(* IEC 61131-3 sources: traffic-lights/PLC_TrafficLights/Class/Varan_Base (part 2) *)

  ud_timeout := ud_ResponseTimeMax + ud_bytes * VM_TIMEOUT_ONE_BYTE + VM_RETRY_TIMEOUT_STD_OFFSET;

END_FUNCTION // Varan_Base::GetRetryTimeout
//=================================================================================================
//---------------------- Additional functions------------------------------------------------------
//=================================================================================================

//[#ENGLISH]
//=================================================================================================
//Function to Start time measurement
//=================================================================================================
#pragma warning(disable:74)
#pragma warning(disable:73)
FUNCTION Varan_Base::StartTimeMeasurement
  VAR_INPUT
    usMode (EAX) 	: DINT;
  END_VAR
#ifdef VM_CLASS_TIME_MEASUREMENT
  VAR
    tmpTime : ^t_TimeMeasurementVaran;
  END_VAR

  case usMode of

    //-----------------------------------------------------------

    VARANTIME_RT:
      tmpTime := #s_TimeRt;

    //-----------------------------------------------------------

    VARANTIME_RTPOSTSCAN:
      tmpTime := #s_TimeRtPostScan;

    //-----------------------------------------------------------

    VARANTIME_CY:
      tmpTime := #s_TimeCy;

    //-----------------------------------------------------------

  end_case;

  if ( tmpTime^.us_Activate ) then
    tmpTime^.ud_Timemark := VaranIn.GetNsTime();
  end_if;

#endif

END_FUNCTION // Varan_Base::StartTimeMeasurement
//[#ENGLISH]
//=================================================================================================
//Function to Stop time measurement
//=================================================================================================
FUNCTION Varan_Base::StopTimeMeasurement
  VAR_INPUT
    usMode (EAX) 	: DINT;
  END_VAR
#ifdef VM_CLASS_TIME_MEASUREMENT
  VAR
    tmpTime : ^t_TimeMeasurementVaran;
  END_VAR

  case usMode of

    //-----------------------------------------------------------

    VARANTIME_RT:
      tmpTime := #s_TimeRt;

    //-----------------------------------------------------------

    VARANTIME_RTPOSTSCAN:
      tmpTime := #s_TimeRtPostScan;

    //-----------------------------------------------------------

    VARANTIME_CY:
      tmpTime := #s_TimeCy;

    //-----------------------------------------------------------

  end_case;

  if ( tmpTime^.us_Activate ) then

    //get actual time
    tmpTime^.ud_ActualTime := VaranIn.GetNsTime() - tmpTime^.ud_Timemark;

    //look for maximum time
    if ( tmpTime^.ud_ActualTime > tmpTime^.ud_MaximalTime ) then
      tmpTime^.ud_MaximalTime := tmpTime^.ud_ActualTime;
    end_if;

    //look for minimum time
    if ( tmpTime^.ud_ActualTime < tmpTime^.ud_MinimalTime ) then
      tmpTime^.ud_MinimalTime := tmpTime^.ud_ActualTime;
    end_if;

    //look for average time (100000 cycles)
    if ( tmpTime^.ud_AverageCounter = 100000 ) then

      tmpTime^.ud_AverageTime 	:= tmpTime^.ud_AverageSum / tmpTime^.ud_AverageCounter;
      tmpTime^.ud_AverageSum 	:= 0;
      tmpTime^.ud_AverageCounter := 0;

    else
      tmpTime^.ud_AverageSum += ( tmpTime^.ud_ActualTime / 100 );
      tmpTime^.ud_AverageCounter += 1;
    end_if;
  end_if;

#endif

END_FUNCTION // Varan_Base::StopTimeMeasurement
#pragma warning(default:74)
#pragma warning(default:73)

//[#ENGLISH]
//=================================================================================================
//Function to set state of class
//=================================================================================================
//[>sd_error]type of error
FUNCTION VIRTUAL GLOBAL Varan_Base::SetState
  VAR_INPUT
    sd_error		: t_e_VaranErrors;
  END_VAR

  //only set error if class is ok
  if ( State = _ClassOk ) then

    State := sd_error;

  else
    //only eeprom error can be cleared
    if ( State = _EEPromError & sd_error = _ClassOk ) then
      State := sd_error;
    end_if;
  end_if;

END_FUNCTION //VIRTUAL GLOBAL Varan_Base::SetState
//[#ENGLISH]
//=================================================================================================
//Function to disable device
//=================================================================================================
//[<sd_retval]0=ok, -17=Port no link, -30=client disabled, -31=client cant enable, -100 function not available with this os version, other return code of os
FUNCTION VIRTUAL GLOBAL Varan_Base::DisableDevice
  VAR_OUTPUT
    sd_retval	: DINT;
  END_VAR
  VAR
    nodeProperty    : LSL_PROPERTY_VALUE_PAIR;
  END_VAR

  //look if funtion is available with this os version
  if ( _RTOSVersion >= VM_DISABLE_DEVICE_AVAILABLE ) then

    if b_PayloadSupport then
      nodeProperty.udPropertyId    := ND_PROP_CONNECTION_STATE;
      nodeProperty.udPropertyValue := CN_STATE_DISCONNECTED;
      sd_retval := MULTI_VARAN_iSetNodeProperties(  hNodeHandle           := ud_HandleModule
                                                  , udPropertyCount       := 1
                                                  , psPropertyValuePairs  := #nodeProperty);
    else
      //disable device
      sd_retval := VARAN_iSetNodeEnableStatus	( uiManager		:= ud_VaranManagerNr
                          , pucNode		:= p_VaranPosition
                          , uiNodeStatus	:= 0
                          );
    end_if;

    // if there was an error at disabling it was not caused by a disabled previous module
    if	( sd_retval <> VARANMANAGER_OK ) &
        ( sd_retval <> VARANMANAGER_CLIENT_DISABLED ) &
        ( sd_retval <> VARANMANAGER_ADMIN_DOL_EXECUTION_ERROR	) &	//because if device before is disabled, DA can't work
        ( VaranIn.IsDeviceDisabled() = FALSE ) then

      State := _DisableError;

      //Set VaranMaster off
      VaranIn.SetManagerOff( e_error := State );
    end_if;

    //port is disabled
    b_DisableDevice := FALSE;
    ud_DisableTime := ops.tAbsolute;
  else
    b_DisableDevice := FALSE;
    sd_retval := -100;
  end_if;

  // Force end of Cylic Post Init
  if bPostInitNeeded then
    CheckCyclicPostInitFinished(TRUE);
  end_if;

END_FUNCTION // Varan_Base::DisableDevice
//[#ENGLISH]
//=================================================================================================
//Function to enable device
//=================================================================================================
//[<sd_retval]0=ok, 1=device must disabled for more then 200ms, 2=-100 function not available with this os version, -17=Port no link, -30=client disabled, -31=client cant enable, other return code of os
FUNCTION VIRTUAL GLOBAL Varan_Base::EnableDevice
  VAR_OUTPUT
    sd_retval	: DINT;
  END_VAR
  VAR
    nodeProperty    : LSL_PROPERTY_VALUE_PAIR;
  END_VAR

  //look if funtion is available with this os
  if ( _RTOSVersion >= VM_DISABLE_DEVICE_AVAILABLE ) then

    //look if watchdog time is gone
    if ( ( ops.tAbsolute - ud_DisableTime ) < 200ms ) then
      sd_retval := 1;
      return;
    end_if;

    if b_PayloadSupport then
      nodeProperty.udPropertyId    := ND_PROP_CONNECTION_STATE;
      nodeProperty.udPropertyValue := CN_STATE_CONNECTED;
      sd_retval := MULTI_VARAN_iSetNodeProperties(  hNodeHandle           := ud_HandleModule
                                                  , udPropertyCount       := 1
                                                  , psPropertyValuePairs  := #nodeProperty);
    else
      //enable device
      sd_retval := VARAN_iSetNodeEnableStatus	( uiManager		:= ud_VaranManagerNr
                          , pucNode		:= p_VaranPosition
                          , uiNodeStatus	:= 1
                          );
    end_if;

    //look for an error
    if ( sd_retval <> VARANMANAGER_OK ) then
      State := _EnableError;
    end_if;
  else
    sd_retval := 2;
  end_if;

END_FUNCTION // Varan_Base::EnableDevice
//[#ENGLISH]
//=================================================================================================
//Function to set all Data Objects off
//=================================================================================================
FUNCTION VIRTUAL GLOBAL Varan_Base::SetDOsOff

  //in base class we have no DO's

END_FUNCTION // Varan_Base::SetDOsOff
//[#ENGLISH]
//=================================================================================================
//Function to look if class is disabled
//=================================================================================================
//[<b_disabled]TRUE -> Device is disabled
FUNCTION VIRTUAL GLOBAL Varan_Base::IsDeviceDisabled
  VAR_OUTPUT
    b_disabled		: BOOL;
  END_VAR

  if 	( State = _NoHardware
    | State = _HardwareNotRequiredIRQ
    )
  then
    b_disabled := TRUE;
  else
    //look class above
    b_disabled := VaranIn.IsDeviceDisabled();
  end_if;

END_FUNCTION //VIRTUAL GLOBAL Varan_Base::IsDeviceDisabled
//[#ENGLISH]
//=================================================================================================
//Function to set multiple memory read/write options
//=================================================================================================
//[>us_filter]filter of multicast write
//[>us_sequence]sequence number of device
//[<sd_retval]error code
FUNCTION VIRTUAL GLOBAL Varan_Base::SetMultipleSettings
  VAR_INPUT
    us_filter		: USINT;
    us_sequence		: usint;
  END_VAR
  VAR_OUTPUT
    sd_retval		: DINT;
  END_VAR
  VAR
    a_data			: ARRAY[0..10] OF USINT;
  END_VAR

  //look if class is ok
  if ( State = _ClassOk ) then

    us_MulticastFilter 		:= us_filter;
    us_MultipleSequence		:= us_sequence;

    //set data for direct access
    a_data[ 0 ] := us_MulticastFilter;
    a_data[ 3 ] := us_sequence;
    a_data[ 10 ] := 16#6;					//to trigger watchdog only with watchdog command and multiple read/write command

    // Payload Support
    if b_PayloadSupport then
      //write data with direct access
      sd_retval := MULTI_VARAN_iExecuteDirectAccess(  hNodeHandle := ud_HandleModule
                                                    , udCommand   := VARAN_CMD_CONTROL_WRITE
                                                    , udOffset    := VARAN_MULTIPLE_OFFSET
                                                    , udLength    := sizeof(a_data)
                                                    , pusData     := ( #a_data )$^USINT
                                                    , pudErrorInfo:= NIL);
    else
      //write data with direct access
      sd_retval := VARAN_iWriteControlDA	( uiManager		  := ud_VaranManagerNr
                                          , uiAddress		  := DeviceAddress + VARAN_MULTIPLE_OFFSET
                                          , uiLen			    := sizeof(a_data)
                                          , uiRetryTimeout:= GetRetryTimeout( ud_bytes := sizeof(a_data) )
                                          , pvData		    := ( #a_data )$^UDINT
                                          , puiError		  := NIL
                                          );
    end_if;

    //look if an error occurs
    if ( sd_retval <> VARANMANAGER_OK ) then
      State := _MultipleError;
      return;
    end_if;
  end_if;

END_FUNCTION //VIRTUAL GLOBAL Varan_Base::SetMultipleSettings
//[#ENGLISH]
//=================================================================================================
//Function must be overwrite
//=================================================================================================
//[>p_handle]pointer to data object header
//[>p_data_read]pointer to read data
//[>p_data_write]pointer to data write
//[<sd_retval]error code
#pragma warning(disable: 73)
FUNCTION VIRTUAL GLOBAL Varan_Base::SetMultipleDataPointers
  VAR_INPUT
    p_handle		: ^LSL_VARANFRAME;
    p_data_read		: ^UDINT;
    p_data_write	: ^UDINT;
    DOIndex         : UDINT;
  END_VAR
  VAR_OUTPUT
    sd_retval		: DINT;
  END_VAR

  sd_retval := -1;

END_FUNCTION //VIRTUAL GLOBAL Varan_Base::SetMultipleDataPointers
#pragma warning(default: 73)
//[#ENGLISH]
//=================================================================================================
//Function to get pointer to calib data
//=================================================================================================
//[>p_offset]pointer to variable to write offset
//[<sd_retval]errorcode of os
FUNCTION  Varan_Base::GetCalibDataPointer
  VAR_INPUT
    p_offset	: ^UDINT;
  END_VAR
  VAR_OUTPUT
    sd_retval	: DINT;
  END_VAR
  VAR
    a_data			: ARRAY[0..31] OF UDINT;
    i				: UDINT;
  END_VAR

  //read SPI data
  sd_retval := VaranIn.ReadSPIData( p_us_position_info	:= p_VaranPosition
                  , ud_offset				:= 0
                  , ud_length				:= 128 or VM_SPI_IDENT_LIST
                  , p_data				:= ( #a_data )$^USINT
                  );

  //look for an error
  if ( sd_retval <> VARANMANAGER_OK ) then
    State := _SPIError;
    return;
  end_if;

  //look for right Identifier
  if ( a_data[ 0 ] <> 16#12345678 ) then
    State := _SPIError;
    return;
  end_if;

  //look for valid length	(we only read 128 Byte at the moment [16Byte are header])
  if( a_data[ 3 ] > (128 - 16 ) ) then
    State := _SPIError;
    return;
  end_if;

  //search for calib data
  for i := 0 to a_data[ 3 ] / sizeof( UDINT ) do

    //look for calib id in 3rd byte
    if ( ( a_data[ i + 4 ] and 16#FF00_0000 ) = VM_SPI_CALIB_ID ) then
      p_offset^ := a_data[ i + 4 ] and 16#00FF_FFFF;
      return;
    end_if;
  end_for;

  //if no entry is found
  State := _NoCalibDataFound;
  sd_retval := -100;

END_FUNCTION // Varan_Base::GetCalibDataPointer
//[#ENGLISH]
//=================================================================================================
//Function to get pointer to calib data
//=================================================================================================
//[>ud_offset]offset in SPI - Flash
//[>ud_length]length of data
//[>p_data]pointer to allocated data space
//[<sd_retval]return value of OS
FUNCTION  Varan_Base::ReadSPIData
  VAR_INPUT
    ud_offset	: UDINT;
    ud_length	: UDINT;
    p_data		: ^USINT;
  END_VAR
  VAR_OUTPUT
    sd_retval	: DINT;
  END_VAR
  VAR
    ud_read_length	: UDINT;
  END_VAR

  //look if we have a length
  if ( ud_length = 0 ) then
    sd_retval := -100;
    return;
  end_if;

  //look if data is in one page
  while ( ud_length <> 0 ) do

    //if length is above page size
    if ( ( ud_offset and 16#FF ) + ud_length > 16#FF ) then
      //how many bytes are in this page available
      ud_read_length := 16#100 - ( ud_offset and 16#FF );
      //not more than 128 Bytes
      if ( ud_read_length > 128 ) then
        ud_read_length := 128;
      end_if;
    else
      //not more than 128 Bytes
      if ( ud_length > 128 ) then
        ud_read_length := 128;
      else
        ud_read_length := ud_length;
      end_if;
    end_if;

    //read data
    sd_retval := VaranIn.ReadSPIData( p_us_position_info	:= p_VaranPosition
                    , ud_offset				:= ud_offset
                    , ud_length				:= ud_read_length
                    , p_data				:= p_data
                    );
    //look for an error
    if ( sd_retval <> VARANMANAGER_OK ) then
      State := _SPIError;
      return;
    end_if;

    //correct length
    ud_length -= ud_read_length;
    ud_offset += ud_read_length;
    p_data += ud_read_length;
  end_while;

END_FUNCTION // Varan_Base::ReadSPIData

//[#ENGLISH]
//=================================================================================================
//Function to update module retry counter
//=================================================================================================
FUNCTION VIRTUAL GLOBAL Varan_Base::UpdateRetryCounter
  //function must be override
END_FUNCTION //VIRTUAL GLOBAL Varan_Base::UpdateRetryCounter
//[#ENGLISH]
//=================================================================================================
//Function to get varan time
//=================================================================================================
//[<ud_varan_time]varan time
FUNCTION VIRTUAL GLOBAL Varan_Base::GetVaranTime
  VAR_INPUT
    p_ud_IsoStartPoint	: ^UDINT;
  END_VAR
  VAR_OUTPUT
    ud_varan_time		: UDINT;
  END_VAR

  ud_varan_time := VaranIn.GetVaranTime( p_ud_IsoStartPoint );

END_FUNCTION //VIRTUAL GLOBAL Varan_Base::GetVaranTime
//[#ENGLISH]
//=================================================================================================
//Function to disable Device in Rt (because VARAN_iSetNodeEnableStatus must not called in Realtime)
//=================================================================================================
FUNCTION  Varan_Base::DisableDeviceRt
  VAR_OUTPUT
    sd_retval		: DINT;
  END_VAR

  //look if funtion is available with this os version
  if ( _RTOSVersion >= VM_DISABLE_DEVICE_AVAILABLE ) then

      //disable device
    sd_retval := VaranIn.SetDisableDevice( p_us_position_info := p_VaranPosition );

    //check error
      if ( sd_retval = 0 ) then

        //port is disabled
        b_DisableDevice := FALSE;
        ud_DisableTime := ops.tAbsolute;
      end_if;
  else
    b_DisableDevice := FALSE;
    sd_retval := -100;
  end_if;

  // Force end of Cylic Post Init
  if bPostInitNeeded then
    CheckCyclicPostInitFinished(TRUE);
  end_if;

END_FUNCTION // Varan_Base::DisableDeviceRt

FUNCTION Varan_Base::SetNewPllData
  VAR_INPUT
    ud_delay_time 	: UDINT;
    us_divider 	    : USINT;
  END_VAR
  VAR_OUTPUT
    sd_retval 	    : DINT;
  END_VAR
  VAR
    ud_data			    : UDINT;
  END_VAR

  //calculate right register value (Response Time (in 10ns steps) / 2 - constant FPGA delay time
  ud_DeviceDelayTime := ( p_NodeInfo^.uiResponseTime ) / 20 + VM_CONST_FPGA_DELAY + ud_delay_time;

  // Payload support
  if b_PayloadSupport then
    //write Pll time with direct access
    sd_retval := MULTI_VARAN_iExecuteDirectAccess(  hNodeHandle := ud_HandleModule
                                                  , udCommand   := VARAN_CMD_CONTROL_WRITE
                                                  , udOffset    := VARAN_PLL_OFFSET + 16#C
                                                  , udLength    := 3
                                                  , pusData     := ( #ud_DeviceDelayTime )$^USINT
                                                  , pudErrorInfo:= NIL);
  else
    //write Pll time with direct access
    sd_retval := VARAN_iWriteControlDA( uiManager		  := ud_VaranManagerNr
                                      , uiAddress		  := DeviceAddress + VARAN_PLL_OFFSET + 16#C
                                      , uiLen			    := 3
                                      , uiRetryTimeout:= GetRetryTimeout( ud_bytes := 3 )
                                      , pvData		    := ( #ud_DeviceDelayTime )$^UDINT
                                      , puiError		  := NIL
                                      );
  end_if;

  //look if an error occurs
  if ( sd_retval <> VARANMANAGER_OK ) then
    State := _PllError;
    return;
  end_if;

  //set divider (only for new pll if function is available)
  if ( us_divider <> 0 ) then

    if b_PayloadSupport then  //  -------------------------------------------------------------------------
      // disable divider
      ud_data := 0;

      sd_retval := MULTI_VARAN_iExecuteDirectAccess(  hNodeHandle := ud_HandleModule
                                                    , udCommand   := VARAN_CMD_CONTROL_WRITE
                                                    , udOffset    := VARAN_PLL_OFFSET + 16#A
                                                    , udLength    := 1
                                                    , pusData     := ( #ud_data )$^USINT
                                                    , pudErrorInfo:= NIL);

      //look if an error occurs
      if ( sd_retval <> VARANMANAGER_OK ) then
        State := _PllError;
        return;
      end_if;

      // set divider value
      ud_data := us_divider;

      sd_retval := MULTI_VARAN_iExecuteDirectAccess(  hNodeHandle := ud_HandleModule
                                                    , udCommand   := VARAN_CMD_CONTROL_WRITE
                                                    , udOffset    := VARAN_PLL_OFFSET + 16#B
                                                    , udLength    := 1
                                                    , pusData     := ( #ud_data )$^USINT
                                                    , pudErrorInfo:= NIL);

      //look if an error occurs
      if ( sd_retval <> VARANMANAGER_OK ) then
        State := _PllError;
        return;
      end_if;

      // enable divider
      ud_data := 2#10010000;    //Defaultvalue = 0x80 + SyncDivider Eanble Bit (Bit4)

      sd_retval := MULTI_VARAN_iExecuteDirectAccess(  hNodeHandle := ud_HandleModule
                                                    , udCommand   := VARAN_CMD_CONTROL_WRITE
                                                    , udOffset    := VARAN_PLL_OFFSET + 16#A
                                                    , udLength    := 1
                                                    , pusData     := ( #ud_data )$^USINT
                                                    , pudErrorInfo:= NIL);

      //look if an error occurs
      if ( sd_retval <> VARANMANAGER_OK ) then
        State := _PllError;
        return;
      end_if;

    else  // if b_PayloadSupport -------------------------------------------------------------------------

      // disable divider
      ud_data := 0;

      // write control register
      sd_retval := VARAN_iWriteControlDA( uiManager		  := ud_VaranManagerNr
                                        , uiAddress		  := DeviceAddress + VARAN_PLL_OFFSET + 16#A
                                        , uiLen			    := 1
                                        , uiRetryTimeout:= GetRetryTimeout( ud_bytes := 1 )
                                        , pvData		    := ( #ud_data )$^UDINT
                                        , puiError		  := NIL
                                        );

      //look if an error occurs
      if ( sd_retval <> VARANMANAGER_OK ) then
        State := _PllError;
        return;
      end_if;

      // set divider value
      ud_data := us_divider;

      //write Divider with direct access
      sd_retval := VARAN_iWriteControlDA( uiManager		  := ud_VaranManagerNr
                                        , uiAddress		  := DeviceAddress + VARAN_PLL_OFFSET + 16#B
                                        , uiLen			    := 1
                                        , uiRetryTimeout:= GetRetryTimeout( ud_bytes := 1 )
                                        , pvData		    := ( #ud_data )$^UDINT
                                        , puiError		  := NIL
                                        );

      //look if an error occurs
      if ( sd_retval <> VARANMANAGER_OK ) then
        State := _PllError;
        return;
      end_if;

      // enable divider
      ud_data := 2#10010000;    //Defaultvalue = 0x80 + SyncDivider Eanble Bit (Bit4)

      //write Divider with direct access
      sd_retval := VARAN_iWriteControlDA( uiManager		  := ud_VaranManagerNr
                                        , uiAddress		  := DeviceAddress + VARAN_PLL_OFFSET + 16#A
                                        , uiLen			    := 1
                                        , uiRetryTimeout:= GetRetryTimeout( ud_bytes := 1 )
                                        , pvData		    := ( #ud_data )$^UDINT
                                        , puiError		  := NIL
                                        );

      //look if an error occurs
      if ( sd_retval <> VARANMANAGER_OK ) then
        State := _PllError;
        return;
      end_if;

    end_if; // if b_PayloadSupport -------------------------------------------------------------------------

  end_if; // us_divider <> 0

END_FUNCTION

FUNCTION VIRTUAL GLOBAL Varan_Base::GetDocumentation
  VAR_INPUT
    p_dpne 	: ^CHAR;
  END_VAR
  VAR_OUTPUT
    sd_retval 	: DINT;
  END_VAR

  sd_retval := VaranIn.GetDocumentation(p_us_position_info:=p_VaranPosition, p_dpne:=p_dpne);

END_FUNCTION

FUNCTION VIRTUAL GLOBAL Varan_Base::UpdateRtPostScan

END_FUNCTION

FUNCTION GLOBAL Varan_Base::SetRunStatus
  VAR_INPUT
    state 	: USINT;
  END_VAR
  VAR_OUTPUT
    us_retval 	: USINT;
  END_VAR

  if Required then
    us_retval := state or VARAN_DO_REQUIRED;
  else
    us_retval := state;
  end_if;

END_FUNCTION

FUNCTION VIRTUAL GLOBAL Varan_Base::GetPointer2ObjectPath
  VAR_OUTPUT
    p_us_ObjectPath 	: ^USINT;
  END_VAR
  VAR
    i                       : USINT;
    udSystemVaranManagerCnt : UDINT;
    _Para 	                : CmdStruct;
    _Result 	              : Results;
  END_VAR

  if ( p_ObjectPath = NIL ) then

    if ( p_VaranPosition = NIL ) then

      Varan_Base::Init();

      if ( p_VaranPosition = NIL ) then

        p_us_ObjectPath := NIL;
        return;

      end_if;
    end_if;

    if ( p_VaranPosition^ >= VARAN_MAX_DEPTH ) then
      p_us_ObjectPath := NIL;
      return;
    end_if;

    //alloc memory
    p_ObjectPath := ( To_StdLib.Malloc( size := p_VaranPosition^ + 5 ) )$^USINT;

    To_StdLib.MemCpy( dest 		:= p_ObjectPath
                    , source	:= p_VaranPosition
                    , size		:= p_VaranPosition^ + 1
                    );

    _Para.uiCmd := VM_CMD_GET_SYSTEM_MANAGER_CNT;
    _Result.aData[0]$UDINT  := 1;   // Set to 1 in case the NewInst Method is not Implemented
    udSystemVaranManagerCnt := 1;

    if VaranIn.NewInst(#_Para, #_Result) = READY then
      udSystemVaranManagerCnt := _Result.aData[0]$UDINT;
    end_if;

    //Check if we have to build the "new" hardware tree with the new escape sequence
    if udSystemVaranManagerCnt > 1 then

      //More than one manager --> new HW-Tree with new esacpe sequence

      //insert one byte after length
      for i := p_ObjectPath^ to 1 by -1 do
        ( p_ObjectPath + i + 4 )^ := ( p_ObjectPath + i )^;
      end_for;

      // domain info byte
      ( p_ObjectPath + 1 )^ := 0;

      //insert escape sequence for varan
      ( p_ObjectPath + 2 )^ := HWT_ESCAPE_MULTIVARAN;

      //insert escape sequence for varan
      ( p_ObjectPath + 3 )^ := ud_VaranManagerNr$USINT;

      //insert escape sequence for varan
      ( p_ObjectPath + 4 )^ := HWT_ESCAPE_VARAN;

      //increase length
      p_ObjectPath^ += 4;

    else

      //Old HW-Tree (without Multivaran Escape sequence)

      //insert one byte after length
      for i := p_ObjectPath^ to 1 by -1 do
        ( p_ObjectPath + i + 2 )^ := ( p_ObjectPath + i )^;
      end_for;

      // domain info byte
      ( p_ObjectPath + 1 )^ := 0;

      //insert escape sequence for varan
      ( p_ObjectPath + 2 )^ := HWT_ESCAPE_VARAN;

      //increase length
      p_ObjectPath^ += 2;

    end_if;

    //register object path in OS
    SetObjectThisp(p_us_ObjectPath:=p_ObjectPath, ud_thisp:=this$UDINT);

  end_if;

  p_us_ObjectPath := p_ObjectPath;

END_FUNCTION

FUNCTION VIRTUAL GLOBAL Varan_Base::SetObjectThisp
  VAR_INPUT
    p_us_ObjectPath 	: ^USINT;
    ud_thisp 	: UDINT;
  END_VAR
  VAR_OUTPUT
    sd_retval 	: DINT;
  END_VAR

  sd_retval := VaranIn.SetObjectThisp(p_us_ObjectPath,ud_thisp);

END_FUNCTION

FUNCTION VIRTUAL GLOBAL Varan_Base::GetObjectThisp
  VAR_INPUT
    p_us_ObjectPath : ^USINT;
  END_VAR
  VAR_OUTPUT
    ud_Thisp 	      : UDINT;
  END_VAR

  ud_thisp := VaranIn.GetObjectThisp(p_us_ObjectPath:=p_us_ObjectPath);

END_FUNCTION

FUNCTION Varan_Base::Diagnose
#ifdef VARAN_DIAGNOSE
  VAR
    os_retcode : DINT;
  END_VAR

  if State = _ClassOk then
    os_retcode := VARAN_IGETVARANDIAGNOSTICS(8, #s_Diagnose.cmd_Input, s_Diagnose.InputSize, #s_Diagnose.cmd_Output, #s_Diagnose.OutputSize);

    //reset counter
    if s_Diagnose.Command = Reset then
      ConnectCounter      := 0;
      FaultCounter        := 0;
      RXLost              := 0;
      TXLost              := 0;
      s_Diagnose.Command  := Activate;
    end_if;

    //OS doesn't support Diagnose
    if os_retcode <> 0 then
      DiagControl := -1;
      return;
    end_if;

    //FPGA doesn't support Diagnose
    if s_Diagnose.cmd_Output.Flags.1 = 0 then
      DiagControl := -2;
      return;
    end_if;

    DiagControl     := 1;
    ConnectCounter  += s_Diagnose.cmd_Output.Counter1 - s_Diagnose.OldCounter.Counter1;
    FaultCounter    += s_Diagnose.cmd_Output.Counter2 - s_Diagnose.OldCounter.Counter2;
    RXLost          += s_Diagnose.cmd_Output.Counter3 - s_Diagnose.OldCounter.Counter3;
    TXLost          += s_Diagnose.cmd_Output.Counter4 - s_Diagnose.OldCounter.Counter4;

    s_Diagnose.OldCounter.Counter1 := s_Diagnose.cmd_Output.Counter1;
    s_Diagnose.OldCounter.Counter2 := s_Diagnose.cmd_Output.Counter2;
    s_Diagnose.OldCounter.Counter3 := s_Diagnose.cmd_Output.Counter3;
    s_Diagnose.OldCounter.Counter4 := s_Diagnose.cmd_Output.Counter4;
  end_if;
#endif
END_FUNCTION

#pragma warning(disable:73)
#pragma warning(disable:74)
#pragma warning(disable:76)
FUNCTION VIRTUAL GLOBAL Varan_Base::DiagControl::Write
  VAR_INPUT
    input (EAX) 	: DINT;
  END_VAR
  VAR_OUTPUT
    result (EAX) 	: DINT;
  END_VAR

#ifdef VARAN_DIAGNOSE

  if input >= 0 & input <= 2 then
    s_Diagnose.Command$DINT := input;
  end_if;

#endif

END_FUNCTION
#pragma warning(default:73)
#pragma warning(default:74)
#pragma warning(default:76)

FUNCTION VIRTUAL GLOBAL Varan_Base::ValidateSerNo::Write
  VAR_INPUT
    input (EAX) 	: DINT;
  END_VAR
  VAR_OUTPUT
    result (EAX) 	: DINT;
  END_VAR

  result := input;

  if (b_ValidationInProgress = FALSE) & SerNoValidation then

    To_MultiTask.CREATETHREAD(taskfunction0:=#SerNoValidationTask(),
                              priority0:=14,
                              stackSize0:=16#4000,
                              flags0:=MT_TASK_SAVETHIS,
                              parameter0:=this,
                              name0:=#szSerNoStr[0]);

    b_ValidationInProgress := TRUE;
  end_if;

END_FUNCTION

FUNCTION Varan_Base::SerNoValidationTask

  // get length of string
  SerNoHeader.StringLength := _strlen(#szSerNoStr[0]);

  // reserve enough space in ramfile
  if SerNoBackup.SetSize(sizeof(SerNoHeader) + SerNoHeader.StringLength) <> C_OK then
      b_ValidationInProgress := FALSE;
      return;
    end_if;

  // initialize the rest of the header
  SerNoHeader.Version := SERNO_VALIDATION_VERSION;
  SerNoHeader.ZeroByte := 0;

  // write to ramfile
  if (SerNoBackup.SetDataAt((#SerNoHeader)$^USINT, sizeof(SerNoHeader), 0) = C_OK) &
     (SerNoBackup.SetDataAt((#szSerNoStr[0])$^USINT, _strlen(#szSerNoStr[0]), sizeof(SerNoHeader)) = C_OK) then
    // if we had a problem with serial number before
    if State = _InvalidSerialNo then
      // try to reconnect
      Varan_HwConnect(0);
    end_if;

    ValidateSerNo := 1;
  else
    ValidateSerNo := 0;
  end_if;

  b_ValidationInProgress := FALSE;

END_FUNCTION

#pragma warning(disable:73)
FUNCTION VIRTUAL GLOBAL Varan_Base::CheckDeviceID
  VAR_INPUT
    ID2Check 	: UDINT;
  END_VAR
  VAR_OUTPUT
    IsOK 	: BOOL;
  END_VAR
#pragma warning(default:73)

  IsOK := TRUE;

END_FUNCTION

FUNCTION GLOBAL Varan_Base::FlexInit
  VAR
    sd_retval	: DINT;
  END_VAR

  //look for an error
  if ( pVaran = NIL ) then
    State := _NoVaranInterface;
    if Required then
      VaranIn.AllowRequiredError();
    end_if;
    return;
  end_if;

  //-----------------------------------------------------------------------------------------------
  //get Varan position if we have no position yet
  if ( p_VaranPosition = NIL ) then

    //alloc memory to get position
    p_VaranPosition := ( To_StdLib.Malloc( size := VARAN_MAX_DEPTH + 1 ) )$^USINT;
    //look if an error occurs
    if ( p_VaranPosition = NIL ) then
      State := _RootError;
      return;
    end_if;

  else

    //alloc memory for position pointer
    p_VaranPosition := 	( To_StdLib.ReAlloc	( mptr := p_VaranPosition , newsize	:= VARAN_MAX_DEPTH + 1))$^USINT;
    //look if an error occurs
    if ( p_VaranPosition = NIL ) then
      State := _RootError;
      return;
    end_if;

  end_if;

  //set length to 0
  p_VaranPosition^ := 0;

  //get position
  sd_retval := VaranIn.GetVaranPosition( p_us_info := p_VaranPosition );

  //look if an error occurs
  if ( sd_retval <> VARANMANAGER_OK ) then
    State := _RootError;
    return;
  end_if;

  //alloc memory for position pointer
  p_VaranPosition := 	( To_StdLib.ReAlloc	( mptr		:= p_VaranPosition
                      , newsize	:= p_VaranPosition^ + 1
                      )
            )$^USINT;

  //look if an error occurs
  if ( p_VaranPosition = NIL ) then
    State := _RootError;
    return;
  end_if;

  //-----------------------------------------------------------------------------------------------
  //install callback function
  sd_retval := InstallCallbackObject();

  //look if an error occurs
  if ( sd_retval <> VARANMANAGER_OK ) then
    State := _CallBackError;
    return;
  end_if;

END_FUNCTION

FUNCTION GLOBAL Varan_Base::AllowRequiredError

  VaranIn.AllowRequiredError();

END_FUNCTION

FUNCTION GLOBAL Varan_Base::IsTransparent
  VAR_OUTPUT
    isTransparent 	: BOOL;
  END_VAR

  IF TransparentInfo.ClientTransparentRead = FALSE THEN

    Transparent := Transparent.Read();
    IF Transparent | VaranIn.IsTransparent() THEN
      Transparent := 1;
      TransparentInfo.DeviceIsTransparent := TRUE;
      Required := 0;
    END_IF;

    TransparentInfo.ClientTransparentRead := TRUE;

  END_IF;

  isTransparent := TransparentInfo.DeviceIsTransparent;

END_FUNCTION

FUNCTION VIRTUAL GLOBAL Varan_Base::AddRdPayloadDO
  VAR_INPUT
    ud_dol_type 	: UDINT;
    p_ud_handle 	: ^UDINT;
    ud_offset_read 	: UDINT;
    ud_length_read 	: UDINT;
    p_ud_data_read 	: ^UDINT;
    ud_type 	: UDINT;
    ud_priority 	: UDINT;
    ud_WritePayloadType   : UDINT;
  END_VAR
  VAR_OUTPUT
    sd_retval 	: DINT;
  END_VAR
  VAR
      // For NewInst command
    _Para 	        : CmdStruct;
    _Result 	      : Results;
    paraAddDO       : t_VM_CMD_AddDO;
    paraGetPointers : t_VM_CMD_GetDataPointers;
    dummy           : UDINT;
  END_VAR

  // Add DO Command ------------------------------------------------------------------------------------------
  _Para.uiCmd := VM_CMD_ADD_DO;

  if ud_HandleModule then
    paraAddDO.ud_ModuleHandle := ud_HandleModule;
  else
    sd_retval := VM_CMD_ERROR_MODULE_HANDLE;
    return;
  end_if;

  paraAddDO.p_ud_DoHandle   := p_ud_handle;
  paraAddDO.ud_b_DoRequired := Required$UDINT;
  paraAddDO.ud_DolType      := ud_dol_type;
  paraAddDO.ud_OffsetRead   := ud_offset_read;
  paraAddDO.ud_LengthRead   := ud_length_read;
  paraAddDO.ud_OffsetWrite  := 0;
  paraAddDO.ud_LengthWrite  := 0;

  if TimeBase > 0 then
    paraAddDO.ud_PreScalerCounterThreshold   := TimeBase - 1;
  else
    paraAddDO.ud_PreScalerCounterThreshold   := 0;
  end_if;

  paraAddDO.ud_PreScalerCounterStartValue  := 0;

  if ud_priority = VM_PRIORITY_INVALID then
    // paraAddDO.ud_Priority := VM_PRIORITY_READ_DO;  // Only with Timesplit
    paraAddDO.ud_Priority := VM_PRIORITY_DEFAULT;
  else
    paraAddDO.ud_Priority := ud_priority;
  end_if;

  paraAddDO.ud_Filter   := 0;
  paraAddDO.ud_Slices   := 0;

  if ud_WritePayloadType then
    paraAddDO.ud_WritePayloadType := WR_PLD_TYPE_RD_ACCESS_CONFIGURABLE;
  else
    paraAddDO.ud_WritePayloadType := WR_PLD_TYPE_STANDARD;
  end_if;

  if ud_type = VM_CONTROL_ACCESS then
    paraAddDO.ud_Command  := VARAN_CMD_CONTROL_READ;
  else
    paraAddDO.ud_Command  := VARAN_CMD_MEMORY_READ;
  end_if;

  _Para.aPara[0]  := (#paraAddDO)$DINT;

  _result.aData[0]$DINT := VM_CMD_OK;

  // Add DO via NewInst
  if VaranIn.NewInst(#_Para, #_Result) <> READY &
     _result.aData[0]$DINT = VM_CMD_OK then
    // If NewInst failed but retcode is still OK
    sd_retval := VM_CMD_ERROR_NEW_INST;
  else
    sd_retval := _result.aData[0]$DINT;
  end_if;

  if sd_retval <> VM_CMD_OK then
    return;
  end_if;

  // Get Pointers Command ------------------------------------------------------------------------------------------
  _Para.uiCmd := VM_CMD_GET_DATA_POINTERS;

  if p_ud_handle^ then
    paraGetPointers.ud_DoHandle     := p_ud_handle^;
  else
    sd_retval := VM_CMD_ERROR_DO_HANDLE;
    return;
  end_if;

  paraGetPointers.p_ud_ReadData   := p_ud_data_read;
  paraGetPointers.p_ud_WriteData  := #dummy;

  _Para.aPara[0]  := (#paraGetPointers)$DINT;
  _result.aData[0]$DINT := VM_CMD_OK;

  // Get Data Poiners via NewInst
  if VaranIn.NewInst(#_Para, #_Result) <> READY &
     _result.aData[0]$DINT = VM_CMD_OK then
    // If NewInst failed but retcode is still OK
    sd_retval := VM_CMD_ERROR_NEW_INST;
  else
    sd_retval := _result.aData[0]$DINT;
  end_if;

END_FUNCTION

FUNCTION VIRTUAL GLOBAL Varan_Base::AddWrPayloadDO
  VAR_INPUT
    ud_dol_type 	: UDINT;
    p_ud_handle 	: ^UDINT;
    ud_offset_write 	: UDINT;
    ud_length_write 	: UDINT;
    p_ud_data_write 	: ^UDINT;
    ud_type 	: UDINT;
    ud_priority 	: UDINT;
    ud_WritePayloadType   : UDINT;
  END_VAR
  VAR_OUTPUT
    sd_retval 	: DINT;
  END_VAR
  VAR
      // For NewInst command
    _Para 	        : CmdStruct;
    _Result 	      : Results;
    paraAddDO       : t_VM_CMD_AddDO;
    paraGetPointers : t_VM_CMD_GetDataPointers;
    dummy           : UDINT;
  END_VAR

  // Add DO Command ------------------------------------------------------------------------------------------
  _Para.uiCmd := VM_CMD_ADD_DO;

  if ud_HandleModule then
    paraAddDO.ud_ModuleHandle := ud_HandleModule;
  else
    sd_retval := VM_CMD_ERROR_MODULE_HANDLE;
    return;
  end_if;

  paraAddDO.p_ud_DoHandle   := p_ud_handle;
  paraAddDO.ud_b_DoRequired := Required$UDINT;
  paraAddDO.ud_DolType      := ud_dol_type;
  paraAddDO.ud_OffsetRead   := 0;
  paraAddDO.ud_LengthRead   := 0;
  paraAddDO.ud_OffsetWrite  := ud_offset_write;
  paraAddDO.ud_LengthWrite  := ud_length_write;

  if TimeBase > 0 then
    paraAddDO.ud_PreScalerCounterThreshold   := TimeBase - 1;
  else
    paraAddDO.ud_PreScalerCounterThreshold   := 0;
  end_if;
  paraAddDO.ud_PreScalerCounterStartValue  := 0;

  if ud_priority = VM_PRIORITY_INVALID then
    // paraAddDO.ud_Priority := VM_PRIORITY_WRITE_DO;  // Only with Timesplit
    paraAddDO.ud_Priority := VM_PRIORITY_DEFAULT;
  else
    paraAddDO.ud_Priority := ud_priority;
  end_if;

  paraAddDO.ud_Filter   := 0;
  paraAddDO.ud_Slices   := 0;

  if ud_WritePayloadType then
    paraAddDO.ud_WritePayloadType := WR_PLD_TYPE_WR_ACCESS_CONFIGURABLE;
  else
    paraAddDO.ud_WritePayloadType := WR_PLD_TYPE_STANDARD;
  end_if;

  if ud_type = VM_CONTROL_ACCESS then
    paraAddDO.ud_Command  := VARAN_CMD_CONTROL_WRITE;
  else
    paraAddDO.ud_Command  := VARAN_CMD_MEMORY_WRITE;
  end_if;

  _Para.aPara[0]  := (#paraAddDO)$DINT;

  _result.aData[0]$DINT := VM_CMD_OK;

  // Add DO via NewInst
  if VaranIn.NewInst(#_Para, #_Result) <> READY &
     _result.aData[0]$DINT = VM_CMD_OK then
    // If NewInst failed but retcode is still OK
    sd_retval := VM_CMD_ERROR_NEW_INST;
  else
    sd_retval := _result.aData[0]$DINT;
  end_if;

  if sd_retval <> VM_CMD_OK then
    return;
  end_if;

  // Get Pointers Command ------------------------------------------------------------------------------------------
  _Para.uiCmd := VM_CMD_GET_DATA_POINTERS;

  if p_ud_handle^ then
    paraGetPointers.ud_DoHandle     := p_ud_handle^;
  else
    sd_retval := VM_CMD_ERROR_DO_HANDLE;
    return;
  end_if;

  paraGetPointers.p_ud_ReadData   := #dummy;
  paraGetPointers.p_ud_WriteData  := p_ud_data_write;

  _Para.aPara[0]  := (#paraGetPointers)$DINT;
  _result.aData[0]$DINT := VM_CMD_OK;

  // Get Data Poiners via NewInst
  if VaranIn.NewInst(#_Para, #_Result) <> READY &
     _result.aData[0]$DINT = VM_CMD_OK then
    // If NewInst failed but retcode is still OK
    sd_retval := VM_CMD_ERROR_NEW_INST;
  else
    sd_retval := _result.aData[0]$DINT;
  end_if;

END_FUNCTION

FUNCTION VIRTUAL GLOBAL Varan_Base::AddRdWrPayloadDO
  VAR_INPUT
    ud_dol_type 	: UDINT;
    p_ud_handle 	: ^UDINT;
    ud_offset_read 	: UDINT;
    ud_length_read 	: UDINT;
    p_ud_data_read 	: ^UDINT;
    ud_offset_write 	: UDINT;
    ud_length_write 	: UDINT;
    p_ud_data_write 	: ^UDINT;
    ud_type 	: UDINT;
    ud_priority 	: UDINT;
    ud_WritePayloadType   : UDINT;
  END_VAR
  VAR_OUTPUT
    sd_retval 	: DINT;
  END_VAR
  VAR
    // For NewInst command
    _Para 	            : CmdStruct;
    _Result 	          : Results;
    paraAddDO           : t_VM_CMD_AddDO;
    paraGetPointers     : t_VM_CMD_GetDataPointers;
  END_VAR

  // Add DO Command ------------------------------------------------------------------------------------------
  _Para.uiCmd := VM_CMD_ADD_DO;

  if ud_HandleModule then
    paraAddDO.ud_ModuleHandle := ud_HandleModule;
  else
    sd_retval := VM_CMD_ERROR_MODULE_HANDLE;
    return;
  end_if;

  paraAddDO.p_ud_DoHandle   := p_ud_handle;
  paraAddDO.ud_b_DoRequired := Required$UDINT;
  paraAddDO.ud_DolType      := ud_dol_type;
  paraAddDO.ud_OffsetRead   := ud_offset_read;
  paraAddDO.ud_LengthRead   := ud_length_read;
  paraAddDO.ud_OffsetWrite  := ud_offset_write;
  paraAddDO.ud_LengthWrite  := ud_length_write;

  if TimeBase > 0 then
    paraAddDO.ud_PreScalerCounterThreshold   := TimeBase - 1;
  else
    paraAddDO.ud_PreScalerCounterThreshold   := 0;
  end_if;
  paraAddDO.ud_PreScalerCounterStartValue  := 0;

  if ud_priority = VM_PRIORITY_INVALID then
    // paraAddDO.ud_Priority := VM_PRIORITY_READ_DO; // Only with Timesplit
    paraAddDO.ud_Priority := VM_PRIORITY_DEFAULT;
  else
    paraAddDO.ud_Priority := ud_priority;
  end_if;

  paraAddDO.ud_Filter   := 0;
  paraAddDO.ud_Slices   := 0;

  if ud_WritePayloadType then
    // Check if only the read or write part of the Payload DO needs to be changed
    if (ud_WritePayloadType = WR_PLD_TYPE_RD_ACCESS_CONFIGURABLE$UDINT) |
       (ud_WritePayloadType = WR_PLD_TYPE_WR_ACCESS_CONFIGURABLE$UDINT) then
      paraAddDO.ud_WritePayloadType := ud_WritePayloadType;
    else
      paraAddDO.ud_WritePayloadType := WR_PLD_TYPE_RW_ACCESS_CONFIGURABLE;
    end_if;
  else
    paraAddDO.ud_WritePayloadType := WR_PLD_TYPE_STANDARD;
  end_if;

  if ud_type = VM_CONTROL_ACCESS then
    paraAddDO.ud_Command  := VARAN_CMD_CONTROL_READ_WRITE;
  else
    paraAddDO.ud_Command  := VARAN_CMD_MEMORY_READ_WRITE;
  end_if;

  _Para.aPara[0]  := (#paraAddDO)$DINT;

  _result.aData[0]$DINT := VM_CMD_OK;

  // Add DO via NewInst
  if VaranIn.NewInst(#_Para, #_Result) <> READY &
     _result.aData[0]$DINT = VM_CMD_OK then
    // If NewInst failed but retcode is still OK
    sd_retval := VM_CMD_ERROR_NEW_INST;
  else
    sd_retval := _result.aData[0]$DINT;
  end_if;

  if sd_retval <> VM_CMD_OK then
    return;
  end_if;

  // Get Pointers Command ------------------------------------------------------------------------------------------
  _Para.uiCmd := VM_CMD_GET_DATA_POINTERS;

  if p_ud_handle^ then
    paraGetPointers.ud_DoHandle     := p_ud_handle^;
  else
    sd_retval := VM_CMD_ERROR_DO_HANDLE;
    return;
  end_if;

  paraGetPointers.p_ud_ReadData   := p_ud_data_read;
  paraGetPointers.p_ud_WriteData  := p_ud_data_write;

  _Para.aPara[0]  := (#paraGetPointers)$DINT;
  _result.aData[0]$DINT := VM_CMD_OK;

  // Get Data Poiners via NewInst
  if VaranIn.NewInst(#_Para, #_Result) <> READY &
     _result.aData[0]$DINT = VM_CMD_OK then
    // If NewInst failed but retcode is still OK
    sd_retval := VM_CMD_ERROR_NEW_INST;
  else
    sd_retval := _result.aData[0]$DINT;
  end_if;

END_FUNCTION

FUNCTION VIRTUAL GLOBAL Varan_Base::AddMovePayloadDO
  VAR_INPUT
    ud_dol_type 	: UDINT;
    p_ud_handle 	: ^UDINT;
    ud_SourceReadDOHandle 	: UDINT;
    ud_SourceReadOffset 	: UDINT;
    ud_DestinationWriteDOHandle 	: UDINT;
    ud_DestinationWriteOffset 	: UDINT;
    ud_LengthMove 	: UDINT;
    ud_Priority 	: UDINT;
  END_VAR
  VAR_OUTPUT
    sd_retval 	: DINT;
  END_VAR
  VAR
      // For NewInst command
    _Para 	            : CmdStruct;
    _Result 	          : Results;
    paraMovDO           : t_VM_CMD_AddMovDo;
  END_VAR

   // Add Move DO Command ------------------------------------------------------------------------------------------
  _Para.uiCmd := VM_CMD_ADD_MOV_DO;

  paraMovDO.p_ud_DoHandle               := p_ud_handle;
  paraMovDO.ud_b_DoRequired             := Required$UDINT;
  paraMovDO.ud_DolType                  := ud_dol_type;
  paraMovDO.ud_SourceReadDoHandle       := ud_SourceReadDOHandle;
  paraMovDO.ud_SourceReadOffset         := ud_SourceReadOffset;
  paraMovDO.ud_DestinationWriteDoHandle := ud_DestinationWriteDOHandle;
  paraMovDO.ud_DestinationWriteOffset   := ud_DestinationWriteOffset;
  paraMovDO.ud_LengthMove               := ud_LengthMove;

  if TimeBase > 0 then
    paraMovDO.ud_PreScalerCounterThreshold   := TimeBase - 1;
  else
    paraMovDO.ud_PreScalerCounterThreshold   := 0;
  end_if;

  paraMovDO.ud_PreScalerCounterStartValue  := 0;

  if ud_priority = VM_PRIORITY_INVALID then
    paraMovDO.ud_Priority := VM_PRIORITY_READ_DO;
  else
    paraMovDO.ud_Priority := ud_priority;
  end_if;

  _Para.aPara[0]  := (#paraMovDO)$DINT;

  _result.aData[0]$DINT := VM_CMD_OK;

  // Add DO via NewInst via NewInst
  if VaranIn.NewInst(#_Para, #_Result) <> READY &
     _result.aData[0]$DINT = VM_CMD_OK then
    // If NewInst failed but retcode is still OK
    sd_retval := VM_CMD_ERROR_NEW_INST;
  else
    sd_retval := _result.aData[0]$DINT;
  end_if;

END_FUNCTION

FUNCTION VIRTUAL GLOBAL Varan_Base::EnableDO
  VAR_INPUT
    ud_DOHandle 	: UDINT;
    ud_bytes 	: UDINT;
  END_VAR
  VAR_OUTPUT
    sd_retval 	: DINT;
  END_VAR

  // LanSte 12.04.2013 09:11 Use IMULTIVARANMANAGER,
  if b_PayloadSupport then
    sd_retval := MULTI_VARAN_iEnableDo(ud_DOHandle);
  else
    if ud_DOHandle then
      ResetDataObject(p_handleDO:=  ud_DOHandle$PLSL_VARANFRAME,
                      us_state  :=  VARAN_DO_CONT_RUN  ,
                      ud_bytes  :=  ud_bytes);

      sd_retval := VARANMANAGER_OK;
    else
      sd_retval := VARANMANAGER_DO_HANDLE_INVALID;
    end_if;
  end_if;

END_FUNCTION

FUNCTION VIRTUAL GLOBAL Varan_Base::DisableDO
	VAR_INPUT
		ud_DOHandle 	: UDINT;
		ud_bytes 	: UDINT;(* := 0 *)
	END_VAR
	VAR_OUTPUT
		sd_retval 	: DINT;
	END_VAR

  // LanSte 12.04.2013 09:11 Use IMULTIVARANMANAGER,
  if b_PayloadSupport then
    sd_retval := MULTI_VARAN_iDisableDo(ud_DOHandle);
  else
    if ud_DOHandle then
      ResetDataObject	( p_handleDO	:= ud_DOHandle$PLSL_VARANFRAME
                      , us_state		:= VARAN_DO_NO_RUN
                      , ud_bytes		:= ud_bytes
                      );
      //ud_DOHandle$PLSL_VARANFRAME^.ucCtrlStat := VARAN_DO_NO_RUN;
      sd_retval := VARANMANAGER_OK;
    else
      sd_retval := VARANMANAGER_DO_HANDLE_INVALID;
    end_if;
  end_if;

END_FUNCTION

FUNCTION VIRTUAL GLOBAL Varan_Base::GetRetryCounter
  VAR_INPUT
    ud_DOHandle 	: UDINT;
  END_VAR
  VAR_OUTPUT
    us_RetryCounter 	: USINT;
  END_VAR
  VAR
    sd_retval 	: DINT;
  END_VAR

   // LanSte 12.04.2013 09:11 Use IMULTIVARANMANAGER,
  if b_PayloadSupport then
    us_RetryCounter := 16#FF;  // Set Value so that we notice a Problem if the Valeu remains unchanged
    sd_retval := MULTI_VARAN_iGetDoProperty(ud_DOHandle, DO_PROP_FAILED_ACCESS_COUNTER, #us_RetryCounter$UDINT);

  else
    if ud_DOHandle then
      us_RetryCounter := ud_DOHandle$PLSL_VARANFRAME^.ucRetryCounter;
      sd_retval := VARANMANAGER_OK;
    else
      sd_retval := VARANMANAGER_DO_HANDLE_INVALID;
    end_if;
  end_if;

END_FUNCTION

FUNCTION VIRTUAL GLOBAL Varan_Base::ChangeDOLengthOffset
  VAR_INPUT
    ud_DOHandle 	: UDINT;
    ud_offset_read 	: UDINT;
    ud_length_read 	: UDINT;
    ud_offset_write 	: UDINT;
    ud_length_write 	: UDINT;
  END_VAR
  VAR_OUTPUT
    sd_retval 	: DINT;
  END_VAR
  VAR
    ud_PropertyCount    : UDINT;
    s_PropertyValuePair : ARRAY [0..4] of LSL_PROPERTY_VALUE_PAIR;
  END_VAR

  if b_PayloadSupport = false then
    sd_retval := VM_CMD_WRONG_OS;
    return;
  end_if;

  ud_PropertyCount := 0;

  if (ud_offset_read <> VM_DO_PROPERTY_INVALID) then

    s_PropertyValuePair[ud_PropertyCount].udPropertyId    := DO_PROP_READ_OFFSET;
    s_PropertyValuePair[ud_PropertyCount].udPropertyValue := ud_offset_read;

    ud_PropertyCount += 1;
  end_if;

  if ud_length_read <> VM_DO_PROPERTY_INVALID then

    s_PropertyValuePair[ud_PropertyCount].udPropertyId    := DO_PROP_READ_LENGTH;
    s_PropertyValuePair[ud_PropertyCount].udPropertyValue := ud_length_read;

    ud_PropertyCount += 1;

  end_if;

  if ud_offset_write <> VM_DO_PROPERTY_INVALID then
    s_PropertyValuePair[ud_PropertyCount].udPropertyId    := DO_PROP_WRITE_OFFSET;
    s_PropertyValuePair[ud_PropertyCount].udPropertyValue := ud_offset_write;

    ud_PropertyCount += 1;
  end_if;

  if ud_length_write <> VM_DO_PROPERTY_INVALID then
    s_PropertyValuePair[ud_PropertyCount].udPropertyId    := DO_PROP_WRITE_LENGTH;
    s_PropertyValuePair[ud_PropertyCount].udPropertyValue := ud_length_write;

    ud_PropertyCount += 1;
  end_if;

  if ud_PropertyCount then
    sd_retval := MULTI_VARAN_iSetDoProperties(ud_DOHandle, ud_PropertyCount, #s_PropertyValuePair[0] );
  else
    // Data undefined
    sd_retval := VM_CMD_ERROR_NO_PROPERTY;
  end_if;

END_FUNCTION

FUNCTION VIRTUAL GLOBAL Varan_Base::ChangeMovDOLengthOffset
  VAR_INPUT
    ud_MovDOHandle 	: UDINT;
    ud_SourceReadDOHandle 	: UDINT;
    ud_SourceReadOffset 	: UDINT;
    ud_DestinationWriteDOHandle 	: UDINT;
    ud_DestinationWriteOffset 	: UDINT;
    ud_LengthMove 	: UDINT;
  END_VAR
  VAR_OUTPUT
    sd_retval 	: DINT;
  END_VAR
  VAR
    ud_PropertyCount    : UDINT;
    s_PropertyValuePair : ARRAY [0..5] of LSL_PROPERTY_VALUE_PAIR;
  END_VAR

  ud_PropertyCount := 0;

  if (ud_sourceReadDOHandle <> VM_DO_PROPERTY_INVALID) then

    s_PropertyValuePair[ud_PropertyCount].udPropertyId    := DO_PROP_SOURCE_READ_DO;
    s_PropertyValuePair[ud_PropertyCount].udPropertyValue := ud_SourceReadDOHandle;

    ud_PropertyCount += 1;
  end_if;

  if (ud_SourceReadOffset <> VM_DO_PROPERTY_INVALID) then

    s_PropertyValuePair[ud_PropertyCount].udPropertyId    := DO_PROP_READ_OFFSET;
    s_PropertyValuePair[ud_PropertyCount].udPropertyValue := ud_SourceReadOffset;

    ud_PropertyCount += 1;
  end_if;

  if (ud_destinationWriteDOHandle <> VM_DO_PROPERTY_INVALID) then

    s_PropertyValuePair[ud_PropertyCount].udPropertyId    := DO_PROP_DESTINATION_WRITE_DO;
    s_PropertyValuePair[ud_PropertyCount].udPropertyValue := ud_DestinationWriteDOHandle;

    ud_PropertyCount += 1;
  end_if;

  if (ud_DestinationWriteOffset <> VM_DO_PROPERTY_INVALID) then

    s_PropertyValuePair[ud_PropertyCount].udPropertyId    := DO_PROP_WRITE_OFFSET;
    s_PropertyValuePair[ud_PropertyCount].udPropertyValue := ud_DestinationWriteOffset;

    ud_PropertyCount += 1;
  end_if;

  if (ud_lengthmove <> VM_DO_PROPERTY_INVALID) then

    s_PropertyValuePair[ud_PropertyCount].udPropertyId    := DO_PROP_MOVE_DATA_LENGTH;
    s_PropertyValuePair[ud_PropertyCount].udPropertyValue := ud_LengthMove;

    ud_PropertyCount += 1;
  end_if;
  if ud_PropertyCount then
    sd_retval := MULTI_VARAN_iSetDoProperties(ud_MovDOHandle, ud_PropertyCount, #s_PropertyValuePair[0] );
  else
    // Data undefined
    sd_retval := VM_CMD_ERROR_NO_PROPERTY;
  end_if;

END_FUNCTION

FUNCTION VIRTUAL GLOBAL Varan_Base::SetPrescaler
  VAR_INPUT
    ud_DOHandle 	: UDINT;
    Prescaler 	: UDINT;
    PrescalerCnt 	: UDINT;
    b_MultipleTimeBase 	: BOOL;
  END_VAR
  VAR_OUTPUT
    sd_retval 	: DINT;
  END_VAR
  VAR
    ud_PropertyCount    : UDINT;
    s_PropertyValuePair : ARRAY [0..1] of LSL_PROPERTY_VALUE_PAIR;
  END_VAR

  ud_PropertyCount := 0;

  s_PropertyValuePair[0].udPropertyId := DO_PROP_PRESCALER_COUNTER_THRESHOLD;
  ud_PropertyCount += 1;

  if b_MultipleTimeBase then

    // Ensure that there is no Multiplication with 0
    if Prescaler & TimeBase > 1 then
      s_PropertyValuePair[0].udPropertyValue := ((Prescaler + 1) * TimeBase) - 1;
    elsif TimeBase > 1 then
      s_PropertyValuePair[0].udPropertyValue := TimeBase-1;
    else
      // No Prescaler and no Timebase
      // Why was this Method called again?
      s_PropertyValuePair[0].udPropertyValue := 0;
    end_if;

  else

    // Set Prescaler
    s_PropertyValuePair[0].udPropertyValue := Prescaler;

    // Set PrescalerCnt (Optional)
    if PrescalerCnt then
      s_PropertyValuePair[1].udPropertyId := DO_PROP_PRESCALER_COUNTER_INIT_VALUE;
      ud_PropertyCount += 1;

      s_PropertyValuePair[1].udPropertyValue := PrescalerCnt;
    end_if;

  end_if;

  sd_retval := MULTI_VARAN_iSetDoProperties(ud_DOHandle, ud_PropertyCount, #s_PropertyValuePair[0] );

END_FUNCTION

FUNCTION VIRTUAL Varan_Base::InstallCallbackObject
  VAR_OUTPUT
    sd_retval 	: DINT;
  END_VAR

  //-----------------------------------------------------------------------------------------------
  // install callback function
  sd_retval := VaranIn.SetObjectCallback( p_us_position_info  := p_VaranPosition
                                        , ud_action_ptr       := ( #Varan_CallBack() )$UDINT
                                        , ud_thisp            := this$UDINT
                                        , sd_required         := Required
                                        );
END_FUNCTION

FUNCTION VIRTUAL GLOBAL Varan_Base::CreateMutex
  VAR_INPUT
    MutexName 	: ^CHAR;
    pThis 	: ^VirtualBase;
  END_VAR
  VAR_OUTPUT
    pv_RetMutex 	: pVoid;
  END_VAR
  VAR
    str_ObjName : array[0..255] of char;
    str_ObjNamePart1 : array[0..VARAN_MUTEX_NAME_MAX_LENGTH-1] of char;
    str_ObjNamePart2 : array[0..VARAN_MUTEX_NAME_END_LENGTH] of char; // +1 for 0 Termination
    str_CombinedName : array[0..VARAN_MUTEX_NAME_MAX_LENGTH-1] of char;
    str_this : array[0..11] of char; // 2 byty %m, 8 byte Address, 1 byte for 0 Termination

    ud_LenObjName  : UDINT;
    ud_LenStr  : UDINT;
    ud_SepLenStr : UDINT;
    ud_LenCombObjName : UDINT;
    ud_LenThis : UDINT;

  END_VAR

  pv_RetMutex := Nil; // Error OS_CILGetv failed

  if pThis = nil then
    pthis := this;
  end_if;

  if (mt_api = nil) then

    if (mt_apiFetch = nil) then

      if(OS_CILGet("LSL_MULTITASK", #mt_apiFetch$void)) THEN
        mt_apiFetch := NIL;
      end_if;

    end_if;

    mt_api := mt_apiFetch;

  end_if;

  if mt_api then

    _memset(dest:=#str_ObjName[0], usByte:=0, cntr:=sizeof(str_ObjName) );
    _memset(dest:=#str_ObjNamePart1[0], usByte:=0, cntr:=sizeof(str_ObjNamePart1) );
    _memset(dest:=#str_ObjNamePart2[0], usByte:=0, cntr:=sizeof(str_ObjNamePart2) );
    _memset(dest:=#str_CombinedName[0], usByte:=0, cntr:=sizeof(str_CombinedName) );
    _memset(dest:=#str_this[0], usByte:=0, cntr:=sizeof(str_this) );

    ud_LenStr := _strlen(MutexName);

    ud_SepLenStr := _strlen(VARAN_STR_MUTEX_NAME_SEPERATOR);
    ud_LenObjName := _GetObjName(pThis:=pthis, pName:=#str_ObjName[0]);

    if (ud_LenStr < VARAN_MUTEX_NAME_MAX_LENGTH) then
      _strcpy(dest:=#str_CombinedName[0], src:=MutexName);
    else
      _strncpy(dest:=#str_CombinedName[0], src:=MutexName, max:=VARAN_MUTEX_NAME_MAX_LENGTH-1);
    end_if;

    if (ud_LenObjName + ud_LenStr) < VARAN_MUTEX_NAME_MAX_LENGTH then
      _strcat(dest:=#str_CombinedName[0], src:=#str_ObjName[0]);
    else
      _strncpy(dest:=#str_ObjNamePart1[0], src:= #str_ObjName[0], max:= VARAN_MUTEX_NAME_MAX_LENGTH - ud_LenStr - ud_SepLenStr - VARAN_MUTEX_NAME_END_LENGTH - 1);    // Copy Beginning of str_ObjName
      _strncpy(dest:=#str_ObjNamePart2[0], src:= #str_ObjName[ud_LenObjName-VARAN_MUTEX_NAME_END_LENGTH-1], max:=VARAN_MUTEX_NAME_END_LENGTH);  // Copy Last MUTEX_NAME_END_LENGTH Char of str_ObjName

      // Put the Mutex String together
      _strcat(dest:=#str_CombinedName[0], src:= #str_ObjNamePart1[0]);
      _strcat(dest:=#str_CombinedName[0], src:= VARAN_STR_MUTEX_NAME_SEPERATOR);
      _strcat(dest:=#str_CombinedName[0], src:= #str_ObjNamePart2[0]);
    end_if;

    pv_RetMutex := OS_MT_CreateSemaphore(MTSEMATYPE_MUTEX, 1, 0, #str_CombinedName[0]);

    if pv_RetMutex = nil then

      // If Create Mutex failed: Insert the this pointer into the string
      ud_LenCombObjName := _strlen(#str_CombinedName[0]);

      str_this[0] := '0';
      str_this[1] := 'x';
      _itoa(udNumber:=pthis$UDINT, pString:=#str_this[2]);
      ud_LenThis  := _strlen(src:=#str_this[0]);

      _strcpy(dest:=#str_CombinedName[ud_LenCombObjName-ud_LenThis], src:=#str_this[0]);

      pv_RetMutex := OS_MT_CreateSemaphore(MTSEMATYPE_MUTEX, 1, 0, #str_CombinedName[0]);

    end_if;

  end_if;

END_FUNCTION

FUNCTION VIRTUAL GLOBAL Varan_Base::MutexStart
  VAR_INPUT
    pMutex 	: pVoid;
  END_VAR

  if(pMutex <> NIL) then
    OS_MT_WAIT(pMutex);
  end_if;

END_FUNCTION

FUNCTION VIRTUAL GLOBAL Varan_Base::MutexStop
  VAR_INPUT
    pMutex 	: pVoid;
  END_VAR

  if(pMutex <> NIL) then
    OS_MT_SIGNAL(pMutex);
  end_if;

END_FUNCTION

FUNCTION VIRTUAL GLOBAL Varan_Base::SingleRunSM
  VAR_INPUT
    p_DOhandle 	: ^UDINT;
    p_b_DOIsRunning 	: ^t_SingleRunState;
  END_VAR

  // xxxxxxxxxxxxxxxxxxxxxxxxxxxxxxxxxxxxxxxxxxxxxxxxxxxxxxxxxxxxxxxxxxxxxxxxxxxxxxxxxxxxxxxxxxxxxxxxxxxxxxxxxxx
  case p_b_DOIsRunning^ of

    SR_STATE_ENABLE_ME :  // DO is not running and start request is set ----------------------------------------
      EnableDO(ud_DOHandle := p_DOhandle^);
      p_b_DOIsRunning^ := SR_STATE_DISABLE_ME;

    SR_STATE_DISABLE_ME : // DO is running and start request is not set ----------------------------------------
      DisableDO(ud_DOHandle:= p_DOhandle^);
      p_b_DOIsRunning^ := SR_STATE_NOTHING;

    SR_STATE_LEAVE_ME_ENABLED : // DO is running and another start request is set ------------------------------
      p_b_DOIsRunning^ := SR_STATE_DISABLE_ME;

  end_case;

END_FUNCTION

FUNCTION VIRTUAL GLOBAL Varan_Base::State::NewInst
  VAR_INPUT
    pPara 	: ^CmdStruct;
    pResult 	: ^Results;
  END_VAR
  VAR_OUTPUT
    ret_code 	: IprStates;
  END_VAR
  VAR
    p_paraGetModuleHandel : ^t_VM_CMD_GetModuleHandle;
    sd_retval             : dint;

    ud_StrSize : UDINT;
    ud_MaxStrSize : UDINT;

  END_VAR

  p_paraGetModuleHandel:= NIL;
  sd_retval            := VARANMANAGER_FATAL_ERROR;

  ud_StrSize    := 0;
  ud_MaxStrSize := 0;

  ret_code := READY;

  CASE pPara^.uiCmd OF
//**********************************************************************************************************************************************************
    VM_CMD_GET_MODULE_HANDLE :
      p_paraGetModuleHandel := (pPara^.aPara[0])$^t_VM_CMD_GetModuleHandle;

      // Check if the passed position string is the same as this class => same module handle
      // For example CDIAS modules behind a CIV
      if (p_paraGetModuleHandel^.p_us_position_info^ = p_VaranPosition^) &  // Lengths of the pos strings are equal
          (_memcmp(ptr1 := p_paraGetModuleHandel^.p_us_position_info+1, ptr2 := p_VaranPosition+1, cntr := p_VaranPosition^) = 0) then  // Contend of the strings are equal

        if ud_HandleModule then // Check if Module handle has been read. May not be read yet because of init order.
          p_paraGetModuleHandel^.p_ud_module_handle^ := ud_HandleModule;
          pResult^.aData[0]$DINT := VM_CMD_OK;
        else
          // Passes on the NewInst command
          ret_code := VaranIn.NewInst(pPara, pResult);

          if pResult^.aData[0]$DINT = VM_CMD_OK &
             ret_code = READY then
            // Safe the Module Handle to this class as well to avoid unnessary OS Calls
            ud_HandleModule := p_paraGetModuleHandel^.p_ud_module_handle^;
          end_if;
          // Else Let calling class deal with the error
        end_if;

      else
        // Passes on the NewInst command
        ret_code := VaranIn.NewInst(pPara, pResult);
      end_if;
//**********************************************************************************************************************************************************
    CMD_GET_HARDWARE_TREE_ENTRY :

      ret_code := ERROR;
      pResult^.aData$t_HWCGetHardwareTreeEntryOut.retcode := _HWC_RETVAL_ERROR;
      pResult^.aData[0]$t_HWCGetHardwareTreeEntryOut.pStr_NextHardewareTreeEntry := NIL;

      // Don't check for State = _ClassOk, method will be used to compare Real HWT with placed classes

      if p_ObjectPath then
        a_HWTEntryStr[0] := p_ObjectPath^$USINT;
        a_HWTEntryStr[1] := 0;
        //a_HWTEntryStr + 2 because first 2 bytes are length, ObjectPath 1st byte is length,
        _memcpy(ptr1:=#a_HWTEntryStr+2, ptr2:=p_ObjectPath+1, cntr:= a_HWTEntryStr[0]);

        pResult^.aData[0]$t_HWCGetHardwareTreeEntryOut.pStr_NextHardewareTreeEntry := #a_HWTEntryStr[0];

        ret_code := READY;
        pResult^.aData$t_HWCGetHardwareTreeEntryOut.retcode := _HWC_RETVAL_OK_HWTSTR_RETURNED;

        // Compare Module string with passed string
        if pPara^.aPara[0]$t_HWCGetHardwareDiagnosisIn.pStr_HardewareTreeEntry then

          if pPara^.aPara[0]$t_HWCGetHardwareDiagnosisIn.pStr_HardewareTreeEntry$^USINT^ =
             pResult^.aData[0]$t_HWCGetHardwareTreeEntryOut.pStr_NextHardewareTreeEntry$^USINT^ then // Compare Length

            if _memcmp( ptr1:= pPara^.aPara[0]$t_HWCGetHardwareDiagnosisIn.pStr_HardewareTreeEntry // Compare Data
                      , ptr2:= pResult^.aData[0]$t_HWCGetHardwareTreeEntryOut.pStr_NextHardewareTreeEntry
                      , cntr:= pResult^.aData[0]$t_HWCGetHardwareTreeEntryOut.pStr_NextHardewareTreeEntry$^USINT^ + 2) = 0 then  // + 2 for 2 Byte Length

              pResult^.aData$t_HWCGetHardwareTreeEntryOut.retcode :=  _HWC_RETVAL_OK_MODULE_FOUND;
            end_if;
          end_if;
        end_if;

      end_if;

//**********************************************************************************************************************************************************
    CMD_GET_HARDWARE_DIAGNOSIS :

//      //search escape sequence, maybe there is a copple module
////      if (ptmpStr+pPara^.aPara[0]$t_HWCGetHardwareDiagnosisIn.us_current_index)^$USINT  = HWT_ESCAPE_VARAN | HWT_ESCAPE_SDIAS | HWT_ESCAPE_CDIAS | HWT_ESCAPE_DIAS  then
//      if (ptmpStr + pPara^.aPara[0]$t_HWCGetHardwareDiagnosisIn.us_current_index)^$USINT  = HWT_ESCAPE_VARAN (*| HWT_ESCAPE_SDIAS | HWT_ESCAPE_CDIAS | HWT_ESCAPE_DIAS*)  then
//        pPara^.aPara[0]$t_HWCGetHardwareDiagnosisIn.us_current_index += 1;
//        //Call SDIAS Manager New Inst
//        ret_code := p_UserCalls.p_Callback^.pSvrChCmd.NewInst(pPara,pResult);
//        return;
//      end_if;

      pResult^.aData$t_HWCGetHardwareDiagnosisOut.retcode := _HWC_RETVAL_ERROR_CLASS_NOT_ONLINE;
      ret_code := ERROR;

      //Return State and Device ID and set retcode ----------------------------------------------------------
      pResult^.aData$t_HWCGetHardwareDiagnosisOut.ClassState := State;
      pResult^.aData$t_HWCGetHardwareDiagnosisOut.ud_DeviceID := GetDeviceID();

      if State = _NoHardware then
        pResult^.aData$t_HWCGetHardwareDiagnosisOut.retcode := _HWC_RETVAL_ERROR_NO_HARDWARE;
      elsif State = _WrongHardware then
        pResult^.aData$t_HWCGetHardwareDiagnosisOut.retcode := _HWC_RETVAL_ERROR_WRONG_HARDWARE;
      elsif State = _NoCalibDataFound then
        pResult^.aData$t_HWCGetHardwareDiagnosisOut.retcode := _HWC_RETVAL_ERROR_NO_CALIB_DATA_FOUND;
      end_if;
      //------------------------------------------------------------------------------------------------------

      if State = _ClassOk then

        // Set Retcodes --------------------------------------------------------------------------------------------
        pResult^.aData$t_HWCGetHardwareDiagnosisOut.retcode := _HWC_RETVAL_OK;
        ret_code := READY;

        //Data which is already in HWK available
        pResult^.aData[0]$t_HWCGetHardwareDiagnosisOut.ud_DeviceID := DeviceID;
        pResult^.aData[0]$t_HWCGetHardwareDiagnosisOut.ud_VendorID := VendorID;

        // Get Serialno -----------------------------------------------------------------------------------------
        pResult^.aData[0]$t_HWCGetHardwareDiagnosisOut.pStr_SerialNo     := #a_SerialNo[0];  // Will be overwritten if this pointer is not equal

        if (this <> p_this) then

          ud_StrSize := SerialNoStr.GetLength() ;
          pResult^.aData[0]$t_HWCGetHardwareDiagnosisOut.pStr_SerialNo     := NIL;

          if ud_StrSize then

            if (ud_StrSize < sizeof(a_SerialNo)) then // < to account for 0 termination
              // Copy complete string
              SerialNoStr.GetDataAt(pData:=#a_SerialNo[0], udSize:=ud_StrSize, udAt:=0);
              a_SerialNo[ud_StrSize] := 0; // 0 termination
            else
              // Copy part string
              SerialNoStr.GetDataAt(pData:=#a_SerialNo[0], udSize:=sizeof(a_SerialNo)-1, udAt:=0);
              a_SerialNo[sizeof(a_SerialNo)-1] := 0; // 0 termination
            end_if;

            pResult^.aData[0]$t_HWCGetHardwareDiagnosisOut.pStr_SerialNo     := #a_SerialNo[0];
          end_if;
        end_if;

        // FPGA Version ----------------------------------------------------------------------------------------------------------
        pResult^.aData[0]$t_HWCGetHardwareDiagnosisOut.hd_FPGAVersion := Release;

        // FW Version --------------------------------------------------------------------------------------------
        GetFWVersion(pData:=#a_FWVersion[0],sizeof(a_FWVersion));
        pResult^.aData$t_HWCGetHardwareDiagnosisOut.pStr_FWVersion := #a_FWVersion[0];

        // Ordering Version ----------------------------------------------------------------------------------------------------------
        pResult^.aData[0]$t_HWCGetHardwareDiagnosisOut.pStr_OrderingNo := (#a_OrderingNoId + sizeof(t_SPI_CalibHeader))$^CHAR;   // Will be overwritten if this pointer is not equal
        if (this <> p_this) then

          sd_retval := GetHWInfoData(p_offset:=#ud_OffestSPI, ud_id:=VM_SPI_ORDERING_NO_ID);
          //look for an error
          if ( sd_retval = VARANMANAGER_OK ) then

            sd_retval := ReadSPIData( ud_offset := ud_OffestSPI
                                    , ud_length	:= sizeof(a_OrderingNoId)
                                    , p_data	:= ( #a_OrderingNoId )$^USINT
                                    );
            //look for an error
            if ( sd_retval = VARANMANAGER_OK ) then

              //t_SPI_CalibHeader ist gleich groß wie der Header von Ordering No Id
              pResult^.aData[0]$t_HWCGetHardwareDiagnosisOut.pStr_OrderingNo := (#a_OrderingNoId + sizeof(t_SPI_CalibHeader))$^CHAR;

              // Null Termination
              ud_StrSize    := a_OrderingNoId[0]$t_SPI_CalibHeader.ud_ListLength;
              ud_MaxStrSize := sizeof(a_OrderingNoId) - sizeof(t_SPI_CalibHeader);

              (pResult^.aData[0]$t_HWCGetHardwareDiagnosisOut.pStr_OrderingNo + ud_MaxStrSize)^ := 0;
              if ud_StrSize < ud_MaxStrSize then
                (pResult^.aData[0]$t_HWCGetHardwareDiagnosisOut.pStr_OrderingNo + ud_StrSize)^ := 0;
              end_if;
            else
              pResult^.aData[0]$t_HWCGetHardwareDiagnosisOut.pStr_OrderingNo := NIL;
// optional, therefore no reason to set the returncode              pResult^.aData$t_HWCGetHardwareDiagnosisOut.retcode := _HWC_RETVAL_ERROR_VARAN_SPI_ACCESS_FAILED;
            end_if;
          else
            pResult^.aData[0]$t_HWCGetHardwareDiagnosisOut.pStr_OrderingNo := NIL;
// optional, therefore no reason to set the returncode            pResult^.aData$t_HWCGetHardwareDiagnosisOut.retcode := _HWC_RETVAL_ERROR_VARAN_SPI_ACCESS_FAILED;
          end_if;
        end_if;

        // Device Name ----------------------------------------------------------------------------------------
        pResult^.aData[0]$t_HWCGetHardwareDiagnosisOut.pStr_DeviceName     := (#a_DeviceName + sizeof(t_SPI_CalibHeader))$^CHAR;  // Will be overwritten if this pointer is not equal

        if (this <> p_this) then
          sd_retval := GetHWInfoData(p_offset:=#ud_OffestSPI, ud_id:=VM_SPI_DEVICE_NAME_ID);
          //look for an error
          if ( sd_retval = VARANMANAGER_OK ) then

            sd_retval := ReadSPIData( ud_offset := ud_OffestSPI
                                    , ud_length	:= sizeof(a_DeviceName)
                                    , p_data	:= ( #a_DeviceName )$^USINT
                                    );

            //look for an error
            if ( sd_retval = VARANMANAGER_OK ) then
              //t_SPI_CalibHeader ist gleich groß wie der Header von spi device name id
              pResult^.aData[0]$t_HWCGetHardwareDiagnosisOut.pStr_DeviceName := (#a_DeviceName + sizeof(t_SPI_CalibHeader))$^CHAR;

              // Null Termination
              ud_StrSize    := a_DeviceName[0]$t_SPI_CalibHeader.ud_ListLength;
              ud_MaxStrSize := sizeof(a_DeviceName) - sizeof(t_SPI_CalibHeader);

              (pResult^.aData[0]$t_HWCGetHardwareDiagnosisOut.pStr_DeviceName + ud_MaxStrSize)^ := 0;
              if ud_StrSize < ud_MaxStrSize then
                (pResult^.aData[0]$t_HWCGetHardwareDiagnosisOut.pStr_DeviceName + ud_StrSize)^ := 0;
              end_if;

            else
              pResult^.aData[0]$t_HWCGetHardwareDiagnosisOut.pStr_DeviceName := NIL;
// optional, therefore no reason to set the returncode              pResult^.aData$t_HWCGetHardwareDiagnosisOut.retcode := _HWC_RETVAL_ERROR_VARAN_SPI_ACCESS_FAILED;
            end_if;
          else
            pResult^.aData[0]$t_HWCGetHardwareDiagnosisOut.pStr_DeviceName := NIL;
// optional, therefore no reason to set the returncode            pResult^.aData$t_HWCGetHardwareDiagnosisOut.retcode := _HWC_RETVAL_ERROR_VARAN_SPI_ACCESS_FAILED;
          end_if;
        end_if;

        // Vendor Name -----------------------------------------------------------------------------------------
        pResult^.aData[0]$t_HWCGetHardwareDiagnosisOut.pStr_VendorName     := (#a_VendorName + sizeof(t_SPI_CalibHeader))$^CHAR;  // Will be overwritten if this pointer is not equal

        if (this <> p_this) then

          sd_retval := GetHWInfoData(p_offset:=#ud_OffestSPI, ud_id:=VM_SPI_VENDOR_NAME_ID);
          //look for an error
          if ( sd_retval = VARANMANAGER_OK ) then

            sd_retval := ReadSPIData( ud_offset := ud_OffestSPI
                                    , ud_length	:= sizeof(a_VendorName)
                                    , p_data	:= ( #a_VendorName )$^USINT
                                    );
            //look for an error
            if ( sd_retval = VARANMANAGER_OK ) then

              //t_SPI_CalibHeader ist gleich groß wie der Header von spi vendor name id
              pResult^.aData[0]$t_HWCGetHardwareDiagnosisOut.pStr_VendorName := (#a_VendorName + sizeof(t_SPI_CalibHeader))$^CHAR;

              // Null Termination
              ud_StrSize    := a_VendorName[0]$t_SPI_CalibHeader.ud_ListLength;
              ud_MaxStrSize := sizeof(a_VendorName) - sizeof(t_SPI_CalibHeader);

              (pResult^.aData[0]$t_HWCGetHardwareDiagnosisOut.pStr_VendorName + ud_MaxStrSize)^ := 0;
              if ud_StrSize < ud_MaxStrSize then
                (pResult^.aData[0]$t_HWCGetHardwareDiagnosisOut.pStr_VendorName + ud_StrSize)^ := 0;
              end_if;

            else
              pResult^.aData[0]$t_HWCGetHardwareDiagnosisOut.pStr_VendorName := NIL;
// optional, therefore no reason to set the returncode              pResult^.aData$t_HWCGetHardwareDiagnosisOut.retcode := _HWC_RETVAL_ERROR_VARAN_SPI_ACCESS_FAILED;
            end_if;
          else
            pResult^.aData[0]$t_HWCGetHardwareDiagnosisOut.pStr_VendorName := NIL;
// optional, therefore no reason to set the returncode            pResult^.aData$t_HWCGetHardwareDiagnosisOut.retcode := _HWC_RETVAL_ERROR_VARAN_SPI_ACCESS_FAILED;

          end_if;
        end_if;

        // Hardware Veriosn and LiceseNo ----------------------------------------------------------------------------------------------
        pResult^.aData[0]$t_HWCGetHardwareDiagnosisOut.ud_LicenseNo := a_IdentList_LicenseNo_HwRev[VARAN_SPI_IDENT_LICENCENO_OFFSET]$UDINT;    // Will be overwritten if this pointer is not equal
        pResult^.aData[0]$t_HWCGetHardwareDiagnosisOut.hd_HWVersion := a_IdentList_LicenseNo_HwRev[VARAN_SPI_IDENT_HARDWAREVER_OFFSET]$UDINT;  // Will be overwritten if this pointer is not equal

        if (this <> p_this) then

          sd_retval := GetHWInfoData(p_offset:=#ud_OffestSPI, ud_id:=VM_SPI_IDENTIFICATION_LIST);

          //look for an error
          if ( sd_retval = VARANMANAGER_OK ) then

            sd_retval := ReadSPIData( ud_offset := ud_OffestSPI
                                    , ud_length	:= sizeof(a_IdentList_LicenseNo_HwRev )
                                    , p_data	:= ( #a_IdentList_LicenseNo_HwRev )$^USINT
                                    );
            //look for an error
            if ( sd_retval = VARANMANAGER_OK ) then
              pResult^.aData[0]$t_HWCGetHardwareDiagnosisOut.ud_LicenseNo := a_IdentList_LicenseNo_HwRev[VARAN_SPI_IDENT_LICENCENO_OFFSET]$UDINT;
              pResult^.aData[0]$t_HWCGetHardwareDiagnosisOut.hd_HWVersion := a_IdentList_LicenseNo_HwRev[VARAN_SPI_IDENT_HARDWAREVER_OFFSET]$UDINT;
            else

              pResult^.aData[0]$t_HWCGetHardwareDiagnosisOut.ud_LicenseNo := 0;
              pResult^.aData[0]$t_HWCGetHardwareDiagnosisOut.hd_HWVersion := 0;
              pResult^.aData$t_HWCGetHardwareDiagnosisOut.retcode := _HWC_RETVAL_ERROR_VARAN_SPI_ACCESS_FAILED; // mandatory entry => set return value
            end_if;
          else

            pResult^.aData[0]$t_HWCGetHardwareDiagnosisOut.ud_LicenseNo := 0;
            pResult^.aData[0]$t_HWCGetHardwareDiagnosisOut.hd_HWVersion := 0;
            pResult^.aData$t_HWCGetHardwareDiagnosisOut.retcode := _HWC_RETVAL_ERROR_VARAN_SPI_ACCESS_FAILED; // mandatory entry => set return value
          end_if;
        end_if;

        p_this := this;  // Safe this pointer, if method is called with for same class that private variables are still valid, don't need to read again

      end_if; // if State = _ClassOk then

//**********************************************************************************************************************************************************
    CMD_POST_INIT_RT_READY :

      // End PostInit if module is online or module has not been found
      if ((Online = 1) | (bOnline = 0)) then
        ret_code := READY;
      else
        ret_code := BUSY;
      end_if;

//**********************************************************************************************************************************************************
    else
      // Passes on the NewInst command
      ret_code := VaranIn.NewInst(pPara, pResult);
  END_CASE;

END_FUNCTION

#pragma warning(disable: 73)
FUNCTION VIRTUAL GLOBAL Varan_Base::Varan_HwSubBusReady
  VAR_INPUT
    ud_data 	: UDINT;
  END_VAR
  VAR_OUTPUT
    sd_retval 	: DINT;
  END_VAR

  sd_retval := VARANMANAGER_OK;

END_FUNCTION
#pragma warning(default: 73)

FUNCTION Varan_Base::GetHWInfoData
	VAR_INPUT
		p_offset 	: ^UDINT;
    ud_id        : UDINT;
	END_VAR
	VAR_OUTPUT
		sd_retval 	: DINT;
	END_VAR

  VAR
    a_data			: ARRAY[0..31] OF UDINT;
    i				: UDINT;
  END_VAR

 //read SPI data
  sd_retval := VaranIn.ReadSPIData( p_us_position_info	:= p_VaranPosition
                  , ud_offset				:= 0
                  , ud_length				:= 128 or VM_SPI_IDENT_LIST
                  , p_data				:= ( #a_data )$^USINT
                  );

  //look for an error
  if ( sd_retval <> VARANMANAGER_OK ) then
    return;
  end_if;

  //look for right Identifier
  if ( a_data[ 0 ] <> 16#12345678 ) then
    return;
  end_if;

  //look for valid length	(we only read 128 Byte at the moment [16Byte are header])
  if( a_data[ 3 ] > (128 - 16 ) ) then
    return;
  end_if;

  //search for input data
  for i := 0 to a_data[ 3 ] / sizeof( UDINT ) do

    //look for input id in 3rd byte
    if ( ( a_data[ i + 4 ] and 16#FF00_0000 ) = ud_id ) then
      p_offset^ := a_data[ i + 4 ] and 16#00FF_FFFF;
      return;
    end_if;
  end_for;

  //if no entry is found
  sd_retval := -100;

END_FUNCTION

FUNCTION VIRTUAL GLOBAL Varan_Base::GetDeviceID
	VAR_OUTPUT
		output 	: UDINT;
	END_VAR
  //Overwrite this method in derived class

 output := HWC_INVALID_DEVICE_ID;

END_FUNCTION

FUNCTION VIRTUAL Varan_Base::GetFWVersion
	VAR_INPUT
		pData 	: ^CHAR;
		length 	: UDINT;
	END_VAR

  //Overwrite in derived Classes
  if pData then
    if Length >= 1 then
      pData^ := 0;    // Set first byte  to 0 termination = invalid string
    end_if;
  end_if;

END_FUNCTION

FUNCTION Varan_Base::GetPllState
	VAR_OUTPUT
		pllstate 	: BSINT;
	END_VAR
  VAR
  	us_data : BSINT;
    sd_retval		: DINT;
  END_VAR

  pllstate := 0;

  if b_PayloadSupport then  //  -------------------------------------------------------------------------
    // get pll state
    us_data := 0;

    sd_retval := MULTI_VARAN_iExecuteDirectAccess(  hNodeHandle := ud_HandleModule
                                                  , udCommand   := VARAN_CMD_CONTROL_READ
                                                  , udOffset    := VARAN_PLL_OFFSET + 16#A
                                                  , udLength    := 1
                                                  , pusData     := ( #us_data )$^USINT
                                                  , pudErrorInfo:= NIL);

    //look if an error occurs
    if ( sd_retval <> VARANMANAGER_OK ) then
      return;
    end_if;

  else  // if b_PayloadSupport -------------------------------------------------------------------------
    // get pll state
    us_data := 0;

    // write control register
    sd_retval := VARAN_iReadControlDA( uiManager		  := ud_VaranManagerNr
                                      , uiAddress		  := DeviceAddress + VARAN_PLL_OFFSET + 16#A
                                      , uiLen			    := 1
                                      , uiRetryTimeout:= GetRetryTimeout( ud_bytes := 1 )
                                      , pvData		    := ( #us_data )$^UDINT
                                      , puiError		  := NIL
                                      );

    //look if an error occurs
    if ( sd_retval <> VARANMANAGER_OK ) then
      return;
    end_if;

  end_if;

#pragma warning(disable:74);
  pllstate.1 := us_data.7; // enabled
  pllstate.2 := us_data.1; // locked
  pllstate.3 := us_data.3; // delay compensated
#pragma warning(default:74);

END_FUNCTION

FUNCTION VIRTUAL GLOBAL Varan_Base::CheckPostInitNeeded
	VAR_INPUT
		pbPostInitSettings 	: ^t_VM_CMD_NEED_POST_INIT_CALL_SETTINGS;
	END_VAR
	VAR_OUTPUT
		PostInitNeeded 	: BOOL;
	END_VAR

  if pbPostInitSettings <> NIL then
    pbPostInitSettings^ := 0;
  end_if;

  PostInitNeeded 	:= FALSE;

END_FUNCTION

FUNCTION VIRTUAL Varan_Base::CheckCyclicPostInitFinished
	VAR_INPUT
		bForcePostInitEnd 	: BOOL;
	END_VAR

  if ((eCycleWork >= _CycleStartIsoDO) | (bOnline = FALSE) | (bForcePostInitEnd)) then
    _ParaBaseCy.uiCmd   := VM_CMD_POST_INIT_FINISHED;
    _ParaBaseCy.aPara[0]:= this$DINT;
    _ParaBaseCy.aPara[1]:= uiBasePostInitHandle;

    if VaranIn.NewInst(pPara:= #_ParaBaseCy, pResult:= #_ResultBaseCy) <> READY then
      LogError("@017D (Varan_Base::CheckCyclicPostInitFinished) Failed to end PostInit.");
    end_if;

    bPostInitNeeded := FALSE;
  end_if;

END_FUNCTION

#pragma warning(disable: 73);
FUNCTION VIRTUAL Varan_Base::LogError
	VAR_INPUT
		e_msg 	: ^CHAR;
	END_VAR

#ifdef HWC_LogError
  HWC_LogError(this, e_msg);
#endif

END_FUNCTION

FUNCTION VIRTUAL Varan_Base::LogValue
	VAR_INPUT
		pString 	: ^CHAR;
		Value 	: UDINT;
		Value2 	: UDINT;(* := 16#FFFFFFFF *)
		Value3 	: UDINT;(* := 16#FFFFFFFF *)
	END_VAR

#ifdef HWC_LogValue3
  HWC_LogValue3(this, pString, Value, Value2, Value3);
#endif

END_FUNCTION
#pragma warning(default: 73);

FUNCTION VIRTUAL Varan_Base::ConvertHwVersion
	VAR_INPUT
		OriginalHwVer 	: HDINT;
	END_VAR
	VAR_OUTPUT
		DisplayedHwVer 	: HDINT;
	END_VAR

  // if it's a sigmatek device
  if VendorID = VM_VENDOR_ID_SIGMATEK then
    // convert the version info to comply with the module print
    DisplayedHwVer := ((OriginalHwVer AND 16#FF000000) SHR 16) OR // high version
                      ((OriginalHwVer AND 16#000F0000) SHR 12) OR // middle version
                       (OriginalHwVer AND 16#0000000F);           // low version
  else
    // use the original
    DisplayedHwVer := OriginalHwVer;
  end_if;

END_FUNCTION

FUNCTION VIRTUAL Varan_Base::GetRequiredWaitTime
	VAR_OUTPUT
		RequiredWaitTime 	: UDINT;
	END_VAR

  RequiredWaitTime := 0;

END_FUNCTION
